(* PLC project HandWritten, plcinfo tests Hand-written 1 *)
(* stored: creationDateTime 2026-10-12T00:00:00 *)

TYPE Range : INT(-10..10);
END_TYPE

TYPE PInt : POINTER TO INT;
END_TYPE

PROGRAM Ladder
  VAR
    a : BOOL;
    b : BOOL;
    c : BOOL;
    d : BOOL;
    start : BOOL;
    done : BOOL;
    stop : BOOL;
    tmr : TON;
  END_VAR
  VAR  (* added by the conversion: wires and edge detectors of the diagram *)
    R_TRIG1 : R_TRIG;
  END_VAR

(* LD diagram, written out as Structured Text *)
(* Motor permissive *)
d := a AND (b OR NOT c);
R_TRIG1(CLK := start);
tmr(IN := R_TRIG1.Q, PT := T#5s);
IF tmr.Q THEN done := TRUE; END_IF;
IF NOT stop THEN JMP End; END_IF;
End:
RETURN;
END_PROGRAM

FUNCTION Calc : INT
  VAR_INPUT
    x : INT;
    enable : BOOL;
  END_VAR

(* FBD diagram, written out as Structured Text *)
Calc := SEL(NOT enable, x + 1, x);
END_FUNCTION

PROGRAM Sequence
  VAR
    go : BOOL;
    left : BOOL;
  END_VAR

INITIAL_STEP Init:
  Fill(P1);
END_STEP
TRANSITION FROM Init TO Right
  := go;
END_TRANSITION
TRANSITION (PRIORITY := 2) FROM Init TO Left
  := left AND NOT go;
END_TRANSITION
STEP Right:
END_STEP
TRANSITION FROM Right TO Init
  := NOT (left);
END_TRANSITION
STEP Left:
END_STEP
TRANSITION FROM Left TO Init
  := go;
END_TRANSITION

ACTION Fill:
level := level + 1;
END_ACTION
END_PROGRAM

CONFIGURATION Config
  RESOURCE Res ON PLC
    VAR_GLOBAL CONSTANT  (* Limits *)
      LIMITS : ARRAY[1..N_MAX] OF LREAL := [1.5, 3(0.0)];
      X0 AT %IX0.0 : BOOL;
    END_VAR
    TASK Fast(INTERVAL := T#1s500ms, PRIORITY := 1);
    TASK Micro(INTERVAL := T#100us, PRIORITY := 2);
    TASK OnEdge(SINGLE := start, PRIORITY := 3);
    PROGRAM inst0 WITH Fast : Ladder;
    PROGRAM inst1 WITH Micro : Sequence;
  END_RESOURCE
END_CONFIGURATION
